// TIA Portal V20 export
DATA_BLOCK "HMI_COM"   // DB2000
{ S7_Optimized_Access := 'FALSE' }
// stored: AutoNumber false
   VAR RETAIN
      Anlagenbeleuchtung_EIN : Bool := TRUE;
      "NOT-HALT_OK" : Bool := TRUE;
      TUERE_OK : Bool := FALSE;
      LICHTVORHANG_OK : Bool := FALSE;
      Grundstellung_Gesamt : Bool := FALSE;
      Dauer_Einzel_Betrieb : Bool := TRUE;
      Antriebe_EIN : Bool := FALSE;
      Antriebe_sind_EIN : Bool := FALSE;
      Stop_nach_Zyklus : Bool := FALSE;
      Stop_nach_Störung : Bool := FALSE;
      Freigabe_Zyklus : Bool := FALSE;
      Ablauf_Aktiv : Bool := FALSE;
      Leerfahren_angewaehlt : Bool := FALSE;
      Leerfahren_laeuft : Bool := FALSE;
      Leerfahren_ende : Bool := FALSE;
      Reset_Schichtzaehler : Bool := FALSE;
      Reset_Auftragszaehler : Bool := FALSE;
      Speichern_Register : Bool := FALSE;
      Richten_Gesamtanlage : Bool := FALSE;
      BM_Anzeige_Nr : Word := 16#0000;
      AmpelStatus : Word := 16#0000;
      BA_Status : Word := 16#0000;
      Einzelschritt { S7_SetPoint := 'True'} : "Stationsvariablen";
      Manuell_Zylinder1 : "Manuell_Zylinder";
      Manuell_Zylinder2 : "Manuell_Zylinder";
      Manuell_Zylinder3 : "Manuell_Zylinder";
      Manuell_Zylinder4 : "Manuell_Zylinder";
      HMI_Achse_Position { S7_SetPoint := 'True'} : "HMI_Achse_Positionen";
      HMI_Achse_Steuerung { S7_SetPoint := 'True'} : "Datentyp_HMI_Achse_Steuerung";
      HMI_Achse_POS_Überschreiben { S7_SetPoint := 'True'} : "HMI_Achse_Positionen_überschreiben";
      Artikelnummer : Array[0..80] of Char;
      Fertigungsauftragsnummer : Array[0..25] of Char;
      Tür_offen : Array[0..15] of Bool;
      Einrichtbetrieb_aktiv : Bool := FALSE;
      Hauptventil_aus_steuern : Bool := FALSE;
      Taktzeit : Array[0..25] of Time;
      Fehlertext_LinMot : String;
      Artikelnummer_String : String;
      Fertigungsauftragsnummer_String : String;
      Reset_Behaelter : UInt;
      "Status Automatik" : Int;
      Artikel_gewechselt : Bool;
      Status_24V_Sicherung : Int;
      "24V_Sicherung_Reset" : Bool;
      "Messwert 1" : Real;
      "Messwert 2" : Real;
      "Messwert 3" : Real;
      Pos4_Trg_Zuführung : Bool;
      Pos4_Zuführung : Int;
      Pos5_Trg_Zuführung : Bool;
      Pos5_Zuführung : Int;
      Pos71_Trg_Zuführung : Bool;
      Pos71_Zuführung : Int;
      Messmittel_ein : Bool;
      Abläufe_Messmittel : Int;
      Messmittel_Rundlauf_ein : Bool;
      Abläufe_Messmittel_Rundlauf : Int;
      "R&R_ein" : Bool;
      DT_takten : Bool;
   END_VAR
BEGIN
   Einzelschritt.Anwahl_Tipp := FALSE;
   Einzelschritt.Status_Anw := TRUE;
   Einzelschritt.Anwahl_GS := FALSE;
   Einzelschritt.Status_GS := FALSE;
   Einzelschritt.Status_Sicher := FALSE;
   Einzelschritt.Tipp_Plus := FALSE;
   Einzelschritt.LEER := FALSE;
   Einzelschritt.Vorhanden := FALSE;
   Einzelschritt.IO := FALSE;
   Einzelschritt.NIO := FALSE;
   Einzelschritt.Reset_Teilestatus := FALSE;
   Einzelschritt.Manu_Freigabe_SK := FALSE;
   Einzelschritt.Richten_lauft := FALSE;
   Einzelschritt.SNr := 0;
   Artikelnummer[0] := '5';
   Artikelnummer[1] := '0';
   Artikelnummer[2] := '2';
   Artikelnummer[3] := '8';
   Artikelnummer[4] := '4';
   Artikelnummer[5] := '5';
   Artikelnummer[6] := '7';
   Artikelnummer[7] := '1';
   Artikelnummer[8] := ' ';
   Artikelnummer[9] := 'B';
   Artikelnummer[10] := 'u';
   Artikelnummer[11] := 'c';
   Artikelnummer[12] := 'h';
   Artikelnummer[13] := 's';
   Artikelnummer[14] := 'e';
   Artikelnummer[15] := ' ';
   Artikelnummer[16] := 'K';
   Artikelnummer[17] := '9';
   Artikelnummer[18..63] := '$00';
   Artikelnummer[64..68] := ' ';
   Artikelnummer[69] := '$00';
   Artikelnummer[70] := ' ';
   Artikelnummer[71] := '$00';
   Artikelnummer[72..80] := ' ';
   Fertigungsauftragsnummer[0] := '1';
   Fertigungsauftragsnummer[1] := '0';
   Fertigungsauftragsnummer[2] := '3';
   Fertigungsauftragsnummer[3..4] := '5';
   Fertigungsauftragsnummer[5] := '9';
   Fertigungsauftragsnummer[6] := '0';
   Fertigungsauftragsnummer[7] := '4';
   Fertigungsauftragsnummer[8..24] := ' ';
   Fertigungsauftragsnummer[25] := '$00';
   Tür_offen[1..8] := FALSE;
END_DATA_BLOCK
